(*
SPDX-FileCopyrightText: c 2026 Oleksandr Tiutyk <trofimich@gmail.com>
SPDX-License-Identifier: MIT
License: https://opensource.org/license/mit
*)

(*!
<summary>Groups dynamic list copying, borrowing, editing, search, sorting and clear cases.</summary>
<description>
Owns the cases, their fixed registration array and any fixtures borrowed by the cases.
Each borrowed fixture is reserved for its case throughout the group lifetime. Use from one task at a stable address.
</description>
*)

{attribute 'no_assign'}
{attribute 'no_explicit_call' := 'do not call this function block directly'}
FUNCTION_BLOCK DynamicListTestGroup EXTENDS TOF_Testing.TestGroup<15>
VAR_STAT
	{attribute 'hide'}
	_ClassName : STRING := __POUNAME();
END_VAR
VAR
	_AppendList : TOF_Collections.List<0>(valueValidator := 0);
	_InsertList : TOF_Collections.List<0>(valueValidator := 0);
	_GetAndSetList : TOF_Collections.List<0>(valueValidator := 0);
	_FindList : TOF_Collections.List<0>(valueValidator := 0);
	_ContainsList : TOF_Collections.List<0>(valueValidator := 0);
	_ContainsGenericList : TOF_Collections.List<0>(valueValidator := 0);
	_RemoveFirstList : TOF_Collections.List<0>(valueValidator := 0);
	_RemoveMatchedList : TOF_Collections.List<0>(valueValidator := 0);
	_RemoveAtList : TOF_Collections.List<0>(valueValidator := 0);
	_SwapList : TOF_Collections.List<0>(valueValidator := 0);
	_AppendGenericList : TOF_Collections.List<0>(valueValidator := 0);
	_InsertGenericList : TOF_Collections.List<0>(valueValidator := 0);
	_GetAndSetGenericList : TOF_Collections.List<0>(valueValidator := 0);

	_Append : ListAppendTest(name := "Append", parent := THIS^, list := _AppendList);
	_Insert : ListInsertTest(name := "Insert", parent := THIS^, list := _InsertList);
	_GetAndSet : ListGetAndSetTest(name := "GetAndSet", parent := THIS^, list := _GetAndSetList);
	_Find : ListFindTest(name := "Find", parent := THIS^, list := _FindList);
	_Contains : ListContainsTest(name := "Contains", parent := THIS^, list := _ContainsList);
	_ContainsGeneric : ListContainsGenericTest(name := "ContainsGeneric", parent := THIS^, list := _ContainsGenericList);
	_RemoveFirst : ListRemoveFirstTest(name := "RemoveFirst", parent := THIS^, list := _RemoveFirstList);
	_RemoveMatched : ListRemoveMatchedTest(name := "RemoveMatched", parent := THIS^, list := _RemoveMatchedList);
	_RemoveAt : ListRemoveAtTest(name := "RemoveAt", parent := THIS^, list := _RemoveAtList);
	_Swap : ListSwapTest(name := "Swap", parent := THIS^, list := _SwapList);
	_Sort : DynamicListSortTest(name := "Sort", parent := THIS^);
	_AppendGeneric : ListAppendGenericTest(name := "AppendGeneric", parent := THIS^, list := _AppendGenericList);
	_InsertGeneric : ListInsertGenericTest(name := "InsertGeneric", parent := THIS^, list := _InsertGenericList);
	_GetAndSetGeneric : ListGetAndSetGenericTest(
		name := "GetAndSetGeneric",
		parent := THIS^,
		list := _GetAndSetGenericList
	);
	_Clear : DynamicListClearTest(name := "Clear", parent := THIS^);

	_Children : ARRAY [0.._ChildCount - 1] OF TOF_Testing.ITestElement :=
	[
		_Append,
		_Insert,
		_GetAndSet,
		_Find,
		_Contains,
		_ContainsGeneric,
		_RemoveFirst,
		_RemoveMatched,
		_RemoveAt,
		_Swap,
		_Sort,
		_AppendGeneric,
		_InsertGeneric,
		_GetAndSetGeneric,
		_Clear
	];
END_VAR

//! <summary>Borrows the fixed child array. Callers must not modify it.</summary>
{attribute 'monitoring' := 'call'}
PROPERTY Children : REFERENCE TO ARRAY [0.._ChildCount - 1] OF TOF_Testing.ITestElement
GET
Children REF= _Children;
END_GET
END_PROPERTY

//! <summary>Borrows the concrete class name. Callers must not modify it.</summary>
{attribute 'monitoring' := 'call'}
PROPERTY ClassName : REFERENCE TO STRING
GET
ClassName REF= _ClassName;
END_GET
END_PROPERTY

//! <summary>Borrows the compiler-initialized namespace name. Callers must not modify it.</summary>
{attribute 'monitoring' := 'call'}
PROPERTY NamespaceName : REFERENCE TO STRING
GET
NamespaceName REF= CurrentNamespace.Name;
END_GET
END_PROPERTY

//! <summary>Reports the concrete instance size in bytes.</summary>
{attribute 'monitoring' := 'call'}
PROPERTY SelfSize : ULINT
GET
SelfSize := XSIZEOF(THIS^);
END_GET
END_PROPERTY

END_FUNCTION_BLOCK

(* stored: Version 1.1.0.1
   POU DynamicListTestGroup: Id {e828e9b1-fc6d-450a-be31-2ea35ddd8125}, SpecialFunc None
   Property Children: Id {2ce7b68d-a606-4550-bf88-c8b969b1cb3d}
   Get Get: Id {e85c5828-d46e-4e23-8f74-5278b509e0ce}
   Property ClassName: Id {8e968db5-3ff6-4f02-84c1-83214cf8f2a2}
   Get Get: Id {50132e57-01fc-4152-b3ea-d059fe82fde7}
   Property NamespaceName: Id {3ecec8dd-7961-45b1-8ef0-12966e78b8c8}
   Get Get: Id {b93c65c7-1bbc-4091-bcc3-fdfccbbc229c}
   Property SelfSize: Id {00be9755-ae4d-447d-b207-5f89db4346e6}
   Get Get: Id {ae0e87ea-8a38-4a8e-90d8-3bf49ad65185} *)
